Staubli VAL3: autoReturn.pjx

--- autoReturn.pjx ---
Parameters version=s8.15.3Cs9_BS3337 stackSize=5000 millimeterUnit=true
Program file=bIsHome.pgx
Program file=getCurMoveID.pgx
Program file=getMotCount.pgx
Program file=logMoveMsgC.pgx
Program file=logMoveMsgJ.pgx
Program file=logMoveMsgL.pgx
Program file=MoveC.pgx
Program file=MoveJ.pgx
Program file=MoveL.pgx
Program file=resetReturnStack.pgx
Program file=returnMove.pgx
Program file=setReferencePos.pgx
Program file=start.pgx
Program file=stop.pgx
Program file=updateJointPos.pgx
Data file=autoReturn.dtx

--- autoReturn.dtx ---
mdesc mNomSpeed
public num nRecIndex
num nMoveIdRec[200]
trsf trToolRec[200]
jointRx jPointRec[200 2]
num nMoveTypeRec[200]
mdesc mReturn = {accel=5, vel=10, decel=5, leave=1, reach=1}
bool bFirstUpdate
mdesc mSpeedRec[200]
jointRx jRefPoint
num nRefDeviate
bool bPushToStack
bool bExact[200]
num nCurrentMoveID
public bool bInterrupt
num nIndex
bool bHaveGetMoveID

--- start.pgx ---
program start()
begin
  //
  waitEndMove()
end

--- bIsHome.pgx ---
program bIsHome(jointRx x_jHome, bool& x_bAtHome)
begin
  //判断当前位置是否为Home点
  x_bAtHome=(abs((herej()-x_jHome))<{4,4,4,4,4,4})
end

--- getCurMoveID.pgx ---
public program getCurMoveID(bool x_bGetMoveId, string x_sType)
  local bool l_bGetMoveId
begin
  l_bGetMoveId=(x_bGetMoveId==true)
  if !l_bGetMoveId
    if(x_sType=="Stop" or x_sType=="Abort" or x_sType=="End") and !bHaveGetMoveID
      nCurrentMoveID=getMoveId()
      bHaveGetMoveID=true
    endIf
    // bInterrupt=true
  else
    bInterrupt=true
  endIf
end

--- getMotCount.pgx ---
public program getMotCount(bool& x_bContain)
  local num l_nI
begin
  x_bContain=false
  for l_nI= 0 to size(nMoveTypeRec)-1
    if nMoveTypeRec[l_nI]!=-1 and nMoveIdRec[l_nI]!=-1
      x_bContain=true
    endIf
  endFor
end

--- logMoveMsgC.pgx ---
program logMoveMsgC(pointRx x_pPoint1, pointRx x_pPoint2, tool x_tTool, mdesc x_mSpeed, num x_nMoveId)
  local string l_sCode
  local bool l_bResult[2]
  local jointRx l_jRef
  local jointRx l_jResult[2]
begin
  //
  if nRecIndex<200
    // c
    if nRecIndex>=1
      l_jRef=jPointRec[nRecIndex-1,1]
    else
      l_jRef=herej()
    endIf
    l_bResult[0]=pointToJoint(x_tTool,l_jRef,x_pPoint1,l_jResult[0])
    l_bResult[1]=pointToJoint(x_tTool,l_jResult[0],x_pPoint2,l_jResult[1])
    //
    if l_bResult[0]==true and l_bResult[1]==true
      setMutex(bPushToStack)
      jPointRec[nRecIndex,0]=l_jResult[0]
      jPointRec[nRecIndex,1]=l_jResult[1]
      trToolRec[nRecIndex]=x_tTool.trsf
      mSpeedRec[nRecIndex]=x_mSpeed
      nMoveIdRec[nRecIndex]=x_nMoveId
      nMoveTypeRec[nRecIndex]=3
      //logMsg("record moveC."+toString("",nMoveIdRec[nRecIndex]))
      nRecIndex=nRecIndex+1
      bPushToStack=false
    else
      // 无关节解
    endIf
  else
    //popUpMsg("记录点数超过容量.")
  endIf

end

--- logMoveMsgJ.pgx ---
program logMoveMsgJ(jointRx x_jPoint, tool x_tTool, mdesc x_mSpeed, num x_nMoveId, bool x_bExact)
  local string l_sCode
begin

  //
  if nRecIndex<200
    // j
    setMutex(bPushToStack)
    jPointRec[nRecIndex,1]=x_jPoint
    trToolRec[nRecIndex]=x_tTool.trsf
    mSpeedRec[nRecIndex]=x_mSpeed
    nMoveIdRec[nRecIndex]=x_nMoveId
    bExact[nRecIndex]=x_bExact
    nMoveTypeRec[nRecIndex]=2
    //logMsg("record moveJ."+toString("",nMoveIdRec[nRecIndex]))
    nRecIndex=nRecIndex+1
    bPushToStack=false
  else
    //popUpMsg("记录点数超过容量.")
  endIf

end

--- logMoveMsgL.pgx ---
program logMoveMsgL(pointRx x_pPoint, tool x_tTool, mdesc x_mSpeed, num x_nMoveId, bool x_bExact)
  local string l_sCode
  local jointRx l_jRef
  local jointRx l_jResult
  local bool l_bResult
begin
  //
  // 走直线or圆弧时，记录目标点位的joint值参考前一个点的joint（如果是第一次记录，参考herej()）
  if nRecIndex<200
    // l
    if nRecIndex>=1
      l_jRef=jPointRec[nRecIndex-1,1]
    else
      l_jRef=herej()
    endIf
    l_bResult=pointToJoint(x_tTool,l_jRef,x_pPoint,l_jResult)
    //
    if l_bResult==true
      setMutex(bPushToStack)
      jPointRec[nRecIndex,1]=l_jResult
      trToolRec[nRecIndex]=x_tTool.trsf
      mSpeedRec[nRecIndex]=x_mSpeed
      nMoveIdRec[nRecIndex]=x_nMoveId
      bExact[nRecIndex]=x_bExact
      nMoveTypeRec[nRecIndex]=1
      //logMsg("record moveL."+toString("",nMoveIdRec[nRecIndex]))
      nRecIndex=nRecIndex+1
      bPushToStack=false
    else
      // 该位置无关节解
    endIf
  else
    //popUpMsg("记录点数超过容量.")
  endIf

end

--- MoveC.pgx ---
public program MoveC(pointRx x_pPoint1, pointRx x_pPoint2, tool x_tTool, mdesc x_mSpeed, num& x_nMoveId)
// // 圆弧运动movec程序
// // 用该程序替代原val3程序中的movec()指令即可
// // 因为原move指令有返回值moveID，所以这里引入一个x_nMoveId，随参考传递出来
begin
  // ---------------------------------------------------------------------------- //
  // 圆弧运动movec程序
  // 用该程序替代原val3程序中的movec()指令即可
  // 因为原move指令有返回值moveID，所以这里引入一个x_nMoveId，随参考传递出来
  // ---------------------------------------------------------------------------- //
  //
  //
  x_nMoveId=movec(x_pPoint1,x_pPoint2,x_tTool,x_mSpeed)
  // log
  call logMoveMsgC(x_pPoint1,x_pPoint2,x_tTool,x_mSpeed,x_nMoveId)

end

--- MoveJ.pgx ---
public program MoveJ(jointRx x_jPoint, tool x_tTool, mdesc x_mSpeed, num& x_nMoveId, bool x_bExact)
// // 关节运动movej程序
// // 用该程序替代原val3程序中的movej()指令即可
// // 因为原move指令有返回值moveID，所以这里引入一个x_nMoveId，随参考传递出来
  local bool l_bResult
begin
  // ---------------------------------------------------------------------------- //
  // 关节运动movej程序
  // 用该程序替代原val3程序中的movej()指令即可
  // 因为原move指令有返回值moveID，所以这里引入一个x_nMoveId，随参考传递出来
  // ---------------------------------------------------------------------------- //
  //
  //
  l_bResult=isInRange(x_jPoint)
  if l_bResult==true
    x_nMoveId=movej(x_jPoint,x_tTool,x_mSpeed)
    if x_bExact
      waitEndMove()
    endIf
    // log
    call logMoveMsgJ(x_jPoint,x_tTool,x_mSpeed,x_nMoveId,x_bExact)
  else
    // 关节点位超限
  endIf

end

--- MoveL.pgx ---
public program MoveL(pointRx x_pPoint, tool x_tTool, mdesc x_mSpeed, num& x_nMoveId, bool x_bExact)
// // 直线运动movel程序
// // 用该程序替代原val3程序中的movel()指令即可
// // 因为原move指令有返回值moveID，所以这里引入一个x_nMoveId，随参考传递出来
begin
  // ---------------------------------------------------------------------------- //
  // 直线运动movel程序
  // 用该程序替代原val3程序中的movel()指令即可
  // 因为原move指令有返回值moveID，所以这里引入一个x_nMoveId，随参考传递出来
  // ---------------------------------------------------------------------------- //
  //
  //
  //
  // 2023.03.15 pointToJoint()时，l_jRef应该取当前指令的前一个点而不是herej()，否则l_jResult可能出现错的解
  // 解决方法：1.新开一个任务，监控当前moveid，当监控开始执行该点轨迹时，重新pointToJoint()，得到l_jResult（待更新）
  x_nMoveId=movel(x_pPoint,x_tTool,x_mSpeed)
  if x_bExact
    //判断是否精确到达
    waitEndMove()
  endIf
  // log
  call logMoveMsgL(x_pPoint,x_tTool,x_mSpeed,x_nMoveId,x_bExact)

end

--- resetReturnStack.pgx ---
public program resetReturnStack(bool x_bRecHere)
// // 清空所有记录堆栈
// // (可选)清空之后是否自动把当前点设为第一个点
  local num l_nI
  local jointRx l_jPos
  local num l_nMoveId
begin
  // ---------------------------------------------------------------------------- //
  // 清空所有记录的堆栈
  // x_bRecHere: 清空之后是否自动记录当前位置作为第一个点
  // ---------------------------------------------------------------------------- //
  //
  for l_nI= 0 to size(nMoveTypeRec)-1
    nMoveTypeRec[l_nI]=-1
    nMoveIdRec[l_nI]=-1
  endFor
  nRecIndex=0
  nCurrentMoveID=0
  bHaveGetMoveID=false

  // 是否记录当前位置为第一个点
  if x_bRecHere
    l_jPos=herej()
    call MoveJ(l_jPos,flange,mNomSpeed,l_nMoveId,false)
    waitEndMove()
  endIf

end

--- returnMove.pgx ---
public program returnMove(bool x_bToRefOnly, jointRx x_jHome, bool& x_bGetMovId)
// // 开始执行回退运动
  local num l_nCurrMoveId
  local bool l_bResult
  local num l_nI
  local jointRx l_jPos
  local num l_nJ
  local tool l_tTool
  local pointRx l_pPos[5]
  local num l_nEndIndex
  local bool l_bAtHome
begin
  // ---------------------------------------------------------------------------- //
  // 开始执行回退运动
  // 2023.03.16 新增x_bToRefOnly，是否回到参考点即结束
  //x_jHome 机器人Home点
  // ---------------------------------------------------------------------------- //
  // 只有在机器人停止状态下，才能执行
  x_bGetMovId=false
  if isSettled()
    // 1.获取当前moveid
    if !bInterrupt
      //l_nCurrMoveId=getMoveId()
      //nCurrentMoveID=l_nCurrMoveId
      x_bGetMovId=true
      l_nCurrMoveId=nCurrentMoveID
      resetMotion()
    else
      l_nCurrMoveId=nCurrentMoveID
    endIf
    logMsg("Current move ID="+toString(".3",l_nCurrMoveId))
    // 当只记录过点个数<=1时，或运动还没到第一个点时，无法执行回退动作
    // 注：如果需要自动回到初始点，在resetReturnStack()之后，先MoveJ(herej())记录第一个点即可
    if nMoveTypeRec[1]!=-1 or l_nCurrMoveId<=nMoveIdRec[0]
      // 2.和堆栈中的moveid比较，找到介于哪两个点之间
      l_bResult=false
      l_nI=-1
      do
        l_nI=l_nI+1
        if(nMoveIdRec[l_nI]+1>=l_nCurrMoveId) and (nMoveTypeRec>0)
          l_bResult=true
        endIf
      until l_bResult==true or l_nI>=size(nMoveTypeRec)-1
      //
      if l_bResult==true
        logMsg("Find current trajectory index:("+toString("",l_nI-1)+" to "+toString("",l_nI)+"]")
        // moveId正在处于(nMoveIdRec[l_nI-1]和nMoveIdRec[l_nI]]之间
        // 3.回退，先move here，然后第一个点从[l_nI-1]开始
        // 3.1 move here first
        wait(isPowered())
        delay(0.5)
        link(l_tTool,flange)
        //resetMotion()
        l_jPos=herej()
        movej(l_jPos,flange,mReturn)
        waitEndMove()
        // 2023.03.16 判断是否回到ref就结束，寻找堆栈里是否有ref点
        l_nEndIndex=-1
        if x_bToRefOnly==true
          for l_nJ=0 to l_nI-1
            if abs(jPointRec[l_nJ,1]-jRefPoint)<{nRefDeviate,nRefDeviate,nRefDeviate,nRefDeviate,nRefDeviate,nRefDeviate}
              l_nEndIndex=l_nJ
            endIf
          endFor
          if l_nEndIndex<0
            popUpMsg("Can't find reference point in stack, end this program.")
            return
          endIf
        else
          // 直接运动到堆栈的第一个点
          l_nEndIndex=1
        endIf
        //
        // 3.2 判断一个[l_nI-1]到[l_nI]这段轨迹的运动类型，倒走到前一个点[l_nI-1]
        //        for l_nJ=l_nI to l_nEndIndex step -1
        if bInterrupt
          //bInterrupt=false
          l_nJ=nIndex
        else
          l_nJ=l_nI
        endIf
        do
          l_tTool.trsf=trToolRec[l_nJ]
          // 得到基于当前参考joint的正确joint位置
          //          if l_nJ==l_nI
          //            // 回退的第一个点，是基于当前位置的joint
          //            bFirstUpdate=true
          //          else
          //            bFirstUpdate=false
          //          endIf
          //          call updateJointPos(l_nJ-1)
          //
          if nMoveTypeRec[l_nJ]==1
            // movel
            // 往回直线运动，点位是[l_nJ-1]的数据，其他诸如工具都应该是[l_nJ]的数据
            l_pPos=jointToPoint(l_tTool,world,jPointRec[l_nJ-1,1])
            //movel(l_pPos,l_tTool,mSpeedRec[l_nJ])
            movel(l_pPos,l_tTool,mReturn)
            //if bExact[l_nJ-1]
            nIndex=l_nJ
            waitEndMove()
            nIndex=l_nJ-1
            call bIsHome(x_jHome,l_bAtHome)
            //endIf
          elseIf nMoveTypeRec[l_nJ]==2
            // movej
            //movej(jPointRec[l_nJ-1,1],l_tTool,mSpeedRec[l_nJ])
            movej(jPointRec[l_nJ-1,1],l_tTool,mReturn)
            //if bExact[l_nJ-1]
            nIndex=l_nJ
            waitEndMove()
            nIndex=l_nJ-1
            call bIsHome(x_jHome,l_bAtHome)
            //endIf
          elseIf nMoveTypeRec[l_nJ]==3
            // movec
            // find middle point
            link(l_pPos[0],world)
            link(l_pPos[1],world)
            link(l_pPos[2],world)
            l_pPos[0]=jointToPoint(l_tTool,world,jPointRec[l_nJ-1,1])
            l_pPos[1]=jointToPoint(l_tTool,world,jPointRec[l_nJ,0])
            l_pPos[2]=jointToPoint(l_tTool,world,jPointRec[l_nJ,1])
            link(l_pPos[3],world)
            if l_nJ==l_nI
              l_pPos[3].trsf=interpolateC(l_pPos[0].trsf,l_pPos[1].trsf,l_pPos[2].trsf,sel((l_nCurrMoveId-roundDown(l_nCurrMoveId))==0,1,l_nCurrMoveId-roundDown(l_nCurrMoveId))/2)
              movec(l_pPos[3],l_pPos[0],l_tTool,mSpeedRec[l_nJ])
            else
              //l_pPos[3].trsf=interpolateC(l_pPos[0].trsf,l_pPos[1].trsf,l_pPos[2].trsf,0.5)
              movec(l_pPos[1],l_pPos[0],l_tTool,mSpeedRec[l_nJ])
            endIf
            //

          endIf
          l_nJ=l_nJ-1
          //endFor
        until(l_nJ==l_nEndIndex-1 or l_bAtHome)
        //
        waitEndMove()
        wait(isSettled())
        // ---- 这里是否需要resetMotion()？待斟酌
        //resetMotion()
        bInterrupt=false
        logMsg("Auto return finished.")
        x_bGetMovId=false
      endIf
    else
      //
      popUpMsg("Only recorded/move one point or less! Please move to the beginning directly!")
    endIf
  else
    //
    popUpMsg("Robot is moving! Please settled robot first!")
  endIf

end

--- setReferencePos.pgx ---
public program setReferencePos(jointRx x_jPoint, num x_nDeviate)
// // 定义一个参考位置
// // x_jPoint: 设定的参考位置的值
// // x_nDeviate: 相对于reference point，允许的误差
begin
  // ---------------------------------------------------------------------------- //
  // 定义一个参考位置
  // x_jPoint: 设定的参考位置的值
  // x_nDeviate: 相对于reference point，允许的误差
  // ---------------------------------------------------------------------------- //
  jRefPoint=x_jPoint
  nRefDeviate=x_nDeviate
end

--- stop.pgx ---
program stop()
begin
end

--- updateJointPos.pgx ---
program updateJointPos(num x_nIndex)
  local jointRx l_jRef
  local pointRx l_pPos
  local tool l_tTool
  local jointRx l_jResult
begin
  // 回退前，基于后一个点[x_nIndex+1]或当前位置，重新更新jPointRec[x_nIndex]
  if bFirstUpdate==true
    l_jRef=herej()
  else
    // 参考关节l_jRef选择[x_nIndex+1]点
    if nMoveTypeRec[x_nIndex+1]==3
      l_jRef=jPointRec[x_nIndex+1,0]
    else
      l_jRef=jPointRec[x_nIndex+1,1]
    endIf
  endIf
  //
  // update joint
  link(l_tTool,flange)
  l_tTool.trsf=trToolRec[x_nIndex]
  l_pPos=jointToPoint(l_tTool,world,jPointRec[x_nIndex,1])
  pointToJoint(l_tTool,l_jRef,l_pPos,l_jResult)
  if jPointRec[x_nIndex,1]!=l_jResult
    jPointRec[x_nIndex,1]=l_jResult
    logMsg("更新jPointRec["+toString("",x_nIndex)+",1]")
  endIf
  // Movec have two points
  if nMoveTypeRec[x_nIndex]==3
    l_pPos=jointToPoint(l_tTool,world,jPointRec[x_nIndex,0])
    pointToJoint(l_tTool,jPointRec[x_nIndex,1],l_pPos,l_jResult)
    if jPointRec[x_nIndex,0]!=l_jResult
      jPointRec[x_nIndex,0]=l_jResult
      logMsg("更新jPointRec["+toString("",x_nIndex)+",0]")
    endIf
  endIf
end
